Fanuc KAREL source: kc00007.KL

-- PROVISIONAL review KL for V940-1; original PC SHA256 2731dfff6493bfe6b0b3f01bd7a378c67acb8d0421391586f6a4988ddc52f68d
-- Incomplete behavior may be omitted. Consult companion uncertainty JSON. Do not deploy.
PROGRAM KC00007
%NOLOCKGROUP
BEGIN
  -- V9_ZERO_TABLE_METADATA_HINT layout=0002_ascii; no indexed target words; source/name/runtime held
  -- UNRESOLVED_PC offsets 5-51; opcodes 27,22,1C,22,22,22,1C,22,31
  -- UNRESOLVED_PC offsets 56-60; opcodes 7F
END KC00007
